(* IEC 61131-3 sources: plcrex/tests/st_examples, 88 files *)

(* ---- TC003.st ---- *)
// ********************************************************************************
// Program Organization Units: FUNCTION
// ********************************************************************************

FUNCTION TC003
  VAR_OUTPUT
    x1 : BOOL;
  END_VAR

  x1 := TRUE;
END_FUNCTION

(* ---- TC004.st ---- *)
// ********************************************************************************
// Program Organization Units: FUNCTION : DATATYPE
// ********************************************************************************

FUNCTION TC004 : BOOL
    VAR_INPUT
        x1 : BOOL;
    END_VAR
    VAR
        x2: BOOL := FALSE;
    END_VAR

    TC004 := x2;
END_FUNCTION

(* ---- TC005.st ---- *)
// ********************************************************************************
// Program Organization Units: FUNCTION_BLOCK
// ********************************************************************************

FUNCTION_BLOCK TC005
  VAR
    x1 : BOOL;
  END_VAR

  x1:= TRUE;
END_FUNCTION_BLOCK

(* ---- TC006.st ---- *)
// ********************************************************************************
// Variable Declaration List: VAR
// ********************************************************************************

FUNCTION_BLOCK TC006
  VAR
    x1 : BOOL := FALSE;
  END_VAR

  x1:= TRUE;
END_FUNCTION_BLOCK

(* ---- TC006_fbd.st ---- *)
FUNCTION_BLOCK TC006
  VAR_INPUT
    i1 : BOOL;
    i2 : BOOL;
  END_VAR
  VAR_OUTPUT
    o1 : BOOL;
    o2 : BOOL;
    o3 : BOOL;
  END_VAR
  VAR
    l1 : BOOL;
    l2 : TIME := T#5s;
    TON0 : TON;
    AND1_OUT : BOOL;
    XOR3_OUT : BOOL;
    OR13_OUT : BOOL;
  END_VAR

  AND1_OUT := AND(i1, i2);
  TON0(AND1_OUT, l2);
  XOR3_OUT := XOR(AND1_OUT, TON0.Q);
  l1 := XOR3_OUT;
  o1 := TON0.Q;
  o2 := i1;
  OR13_OUT := OR(i2, l1);
  o3 := OR13_OUT;
END_FUNCTION_BLOCK

(* ---- TC007.st ---- *)
// ********************************************************************************
// Interface Declaration List: VAR_INPUT
// ********************************************************************************

FUNCTION_BLOCK TC007
  VAR_INPUT
    x1 : BOOL;
  END_VAR
  VAR
    x2 : BOOL := FALSE;
    x3 : BOOL := FALSE;
  END_VAR

  x2:=x1;
END_FUNCTION_BLOCK

(* ---- TC008.st ---- *)
// ********************************************************************************
// Interface Declaration List: VAR_INPUT
// ********************************************************************************

FUNCTION_BLOCK TC008
  VAR_INPUT
    x1 : BOOL := FALSE;
  END_VAR
  VAR
    x2 : BOOL := FALSE;
    x3 : BOOL := FALSE;
  END_VAR

  x2:=x1;
END_FUNCTION_BLOCK

(* ---- TC009.st ---- *)
// ********************************************************************************
// Interface Declaration List: VAR_OUTPUT
// ********************************************************************************

FUNCTION_BLOCK TC009
  VAR_OUTPUT
    x1 : BOOL;
  END_VAR

  x1 := TRUE;
END_FUNCTION_BLOCK

(* ---- TC010.st ---- *)
// ********************************************************************************
// Interface Declaration List: VAR_OUTPUT
// ********************************************************************************

FUNCTION_BLOCK TC010
  VAR_OUTPUT
    x1 : BOOL := FALSE;
  END_VAR

  x1 := TRUE;
END_FUNCTION_BLOCK

(* ---- TC011.st ---- *)
// ********************************************************************************
// Interface Declaration List: VAR_EXTERNAL
// ********************************************************************************

FUNCTION_BLOCK TC011
  VAR_EXTERNAL
    global : BOOL;
  END_VAR
  VAR
    x1 : BOOL;
  END_VAR

  x1 := global;
END_FUNCTION_BLOCK

(* ---- TC012.st ---- *)
// ********************************************************************************
// Interface Declaration List: VAR_IN_OUT
// ********************************************************************************

FUNCTION_BLOCK TC012
  VAR_IN_OUT
    x1 : BOOL;
  END_VAR

  x1:=TRUE;
END_FUNCTION_BLOCK

(* ---- TC013.st ---- *)
// ********************************************************************************
// Data Types: BOOL
// ********************************************************************************

FUNCTION_BLOCK TC013
  VAR
    x1 : BOOL;
  END_VAR

  x1:=TRUE;
END_FUNCTION_BLOCK

(* ---- TC014.st ---- *)
// ********************************************************************************
// Data Types: INT
// ********************************************************************************

FUNCTION_BLOCK TC014
  VAR
    x1 : INT;
  END_VAR

  x1:=5;
END_FUNCTION_BLOCK

(* ---- TC015.st ---- *)
// ********************************************************************************
// Data Types: DINT
// ********************************************************************************

FUNCTION_BLOCK TC015
  VAR
    x1 : DINT;
  END_VAR

  x1:=5;
END_FUNCTION_BLOCK

(* ---- TC016.st ---- *)
// ********************************************************************************
// Data Types: UINT
// ********************************************************************************

FUNCTION_BLOCK TC016
  VAR
    x1 : UINT;
  END_VAR

  x1:=5;
END_FUNCTION_BLOCK

(* ---- TC017.st ---- *)
// ********************************************************************************
// Data Types: REAL
// ********************************************************************************

FUNCTION_BLOCK TC017
  VAR
    x1 : REAL;
  END_VAR

  x1:=5.0;
END_FUNCTION_BLOCK

(* ---- TC018.st ---- *)
// ********************************************************************************
// Data Types: TIME
// ********************************************************************************

FUNCTION_BLOCK TC018
  VAR
    x1 : TIME;
  END_VAR

  x1:=t#5000ms;
END_FUNCTION_BLOCK

(* ---- TC019.st ---- *)
// ********************************************************************************
// Data Types: ARRAY OF BOOL
// ********************************************************************************

FUNCTION_BLOCK TC019
  VAR
    x1 : ARRAY [1..2] OF BOOL;
  END_VAR

  x1[1]:= TRUE;
END_FUNCTION_BLOCK

(* ---- TC020.st ---- *)
// ********************************************************************************
// Data Types: ARRAY OF INT
// ********************************************************************************

FUNCTION_BLOCK TC020
  VAR
    x1 : ARRAY [1..2] OF INT;
  END_VAR

  x1[1]:= 1;
END_FUNCTION_BLOCK

(* ---- TC021.st ---- *)
// ********************************************************************************
// Data Types: ARRAY OF DINT
// ********************************************************************************

FUNCTION_BLOCK TC021
  VAR
    x1 : ARRAY [1..2] OF DINT;
  END_VAR

  x1[1]:= 1;
END_FUNCTION_BLOCK

(* ---- TC022.st ---- *)
// ********************************************************************************
// Data Types: ARRAY OF UINT
// ********************************************************************************

FUNCTION_BLOCK TC022
  VAR
    x1 : ARRAY [1..2] OF UINT;
  END_VAR

  x1[1]:= 1;
END_FUNCTION_BLOCK

(* ---- TC023.st ---- *)
// ********************************************************************************
// Data Types: ARRAY OF REAL
// ********************************************************************************

FUNCTION_BLOCK TC023
  VAR
    x1 : ARRAY [1..2] OF REAL;
  END_VAR

  x1[1]:= 1.0;
END_FUNCTION_BLOCK

(* ---- TC024.st ---- *)
// ********************************************************************************
// Data Types: ARRAY OF TIME
// ********************************************************************************

FUNCTION_BLOCK TC024
  VAR
    x1 : ARRAY [1..2] OF TIME;
  END_VAR

  x1[1]:= t#5000ms;
END_FUNCTION_BLOCK

(* ---- TC025.st ---- *)
// ********************************************************************************
// Expressions: FALSE
// ********************************************************************************

FUNCTION_BLOCK TC025
  VAR
    x1 : BOOL;
  END_VAR

  x1:=FALSE;
END_FUNCTION_BLOCK

(* ---- TC026.st ---- *)
// ********************************************************************************
// Expressions: TRUE
// ********************************************************************************

FUNCTION_BLOCK TC026
  VAR
    x1 : BOOL;
  END_VAR

  x1:=TRUE;
END_FUNCTION_BLOCK

(* ---- TC027.st ---- *)
// ********************************************************************************
// Expressions: =
// ********************************************************************************

FUNCTION_BLOCK TC027
  VAR
    x1 : INT := 4;
    x2 : INT := 6;
    x3 : BOOL;
  END_VAR

  x3:=x1 = x2;
END_FUNCTION_BLOCK

(* ---- TC028.st ---- *)
// ********************************************************************************
// Expressions: =
// ********************************************************************************

FUNCTION_BLOCK TC028
  VAR
    x1 : INT := 6;
    x2 : INT := 6;
    x3 : BOOL;
  END_VAR

  x3:=x1 = x2;
END_FUNCTION_BLOCK

(* ---- TC029.st ---- *)
// ********************************************************************************
// Expressions: <>
// ********************************************************************************

FUNCTION_BLOCK TC029
  VAR
    x1 : INT := 4;
    x2 : INT := 6;
    x3 : BOOL;
  END_VAR

  x3:=x1 <> x2;
END_FUNCTION_BLOCK

(* ---- TC030.st ---- *)
// ********************************************************************************
// Expressions: <>
// ********************************************************************************

FUNCTION_BLOCK TC030
  VAR
    x1 : INT := 6;
    x2 : INT := 6;
    x3 : BOOL;
  END_VAR

  x3:=x1 <> x2;
END_FUNCTION_BLOCK

(* ---- TC031.st ---- *)
// ********************************************************************************
// Expressions: <
// ********************************************************************************

FUNCTION_BLOCK TC031
  VAR
    x1 : INT := 4;
    x2 : INT := 6;
    x3 : BOOL;
  END_VAR

  x3:=x1 < x2;
END_FUNCTION_BLOCK

(* ---- TC032.st ---- *)
// ********************************************************************************
// Expressions: <
// ********************************************************************************

FUNCTION_BLOCK TC032
  VAR
    x1 : INT := 6;
    x2 : INT := 6;
    x3 : BOOL;
  END_VAR

  x3:=x1 < x2;
END_FUNCTION_BLOCK

(* ---- TC033.st ---- *)
// ********************************************************************************
// Expressions: >
// ********************************************************************************

FUNCTION_BLOCK TC033
  VAR
    x1 : INT := 4;
    x2 : INT := 6;
    x3 : BOOL;
  END_VAR

  x3:=x1 > x2;
END_FUNCTION_BLOCK

(* ---- TC034.st ---- *)
// ********************************************************************************
// Expressions: >
// ********************************************************************************

FUNCTION_BLOCK TC034
  VAR
    x1 : INT := 6;
    x2 : INT := 6;
    x3 : BOOL;
  END_VAR

  x3:=x1 > x2;
END_FUNCTION_BLOCK

(* ---- TC035.st ---- *)
// ********************************************************************************
// Expressions: <=
// ********************************************************************************

FUNCTION_BLOCK TC035
  VAR
    x1 : INT := 4;
    x2 : INT := 6;
    x3 : BOOL;
  END_VAR

  x3:=x1 <= x2;
END_FUNCTION_BLOCK

(* ---- TC036.st ---- *)
// ********************************************************************************
// Expressions: <=
// ********************************************************************************

FUNCTION_BLOCK TC036
  VAR
    x1 : INT := 6;
    x2 : INT := 6;
    x3 : BOOL;
  END_VAR

  x3:=x1 <= x2;
END_FUNCTION_BLOCK

(* ---- TC037.st ---- *)
// ********************************************************************************
// Expressions: >=
// ********************************************************************************

FUNCTION_BLOCK TC037
  VAR
    x1 : INT := 4;
    x2 : INT := 6;
    x3 : BOOL;
  END_VAR

  x3:=x1 >= x2;
END_FUNCTION_BLOCK

(* ---- TC038.st ---- *)
// ********************************************************************************
// Expressions: >=
// ********************************************************************************

FUNCTION_BLOCK TC038
  VAR
    x1 : INT := 6;
    x2 : INT := 6;
    x3 : BOOL;
  END_VAR

  x3:=x1 >= x2;
END_FUNCTION_BLOCK

(* ---- TC039.st ---- *)
// ********************************************************************************
// Expressions: NOT
// ********************************************************************************

FUNCTION_BLOCK TC039
  VAR
    x1 : BOOL := TRUE;
    x2 : BOOL;
  END_VAR

  x1:=NOT x1;
  x2 := TRUE;
END_FUNCTION_BLOCK

(* ---- TC040.st ---- *)
// ********************************************************************************
// Expressions: NOT
// ********************************************************************************

FUNCTION_BLOCK TC040
  VAR
    x1 : BOOL := FALSE;
    x2 : BOOL;
  END_VAR

  x1:=NOT x1;
  x2 := TRUE;
END_FUNCTION_BLOCK

(* ---- TC041.st ---- *)
// ********************************************************************************
// Expressions: AND
// ********************************************************************************

FUNCTION_BLOCK TC041
  VAR
    x1 : BOOL := FALSE;
    x2 : BOOL := FALSE;
	x3 : BOOL;
  END_VAR

  x3:=x1 AND x2;
END_FUNCTION_BLOCK

(* ---- TC042.st ---- *)
// ********************************************************************************
// Expressions: AND
// ********************************************************************************

FUNCTION_BLOCK TC042
  VAR
    x1 : BOOL := TRUE;
    x2 : BOOL := FALSE;
	x3 : BOOL;
  END_VAR

  x3:=x1 AND x2;
END_FUNCTION_BLOCK

(* ---- TC043.st ---- *)
// ********************************************************************************
// Expressions: AND
// ********************************************************************************

FUNCTION_BLOCK TC043
  VAR
    x1 : BOOL := FALSE;
    x2 : BOOL := TRUE;
	x3 : BOOL;
  END_VAR

  x3:=x1 AND x2;
END_FUNCTION_BLOCK

(* ---- TC044.st ---- *)
// ********************************************************************************
// Expressions: AND
// ********************************************************************************

FUNCTION_BLOCK TC044
  VAR
    x1 : BOOL := FALSE;
    x2 : BOOL := TRUE;
	x3 : BOOL;
  END_VAR

  x3:=x1 AND x2;
END_FUNCTION_BLOCK

(* ---- TC045.st ---- *)
// ********************************************************************************
// Expressions: XOR
// ********************************************************************************

FUNCTION_BLOCK TC045
  VAR
    x1 : BOOL := FALSE;
    x2 : BOOL := FALSE;
	x3 : BOOL;
  END_VAR

  x3:=x1 XOR x2;
END_FUNCTION_BLOCK

(* ---- TC046.st ---- *)
// ********************************************************************************
// Expressions: XOR
// ********************************************************************************

FUNCTION_BLOCK TC046
  VAR
    x1 : BOOL := TRUE;
    x2 : BOOL := FALSE;
	x3 : BOOL;
  END_VAR

  x3:=x1 XOR x2;
END_FUNCTION_BLOCK

(* ---- TC047.st ---- *)
// ********************************************************************************
// Expressions: XOR
// ********************************************************************************

FUNCTION_BLOCK TC047
  VAR
    x1 : BOOL := FALSE;
    x2 : BOOL := TRUE;
	x3 : BOOL;
  END_VAR

  x3:=x1 XOR x2;
END_FUNCTION_BLOCK

(* ---- TC048.st ---- *)
// ********************************************************************************
// Expressions: XOR
// ********************************************************************************

FUNCTION_BLOCK TC048
  VAR
    x1 : BOOL := TRUE;
    x2 : BOOL := TRUE;
	x3 : BOOL;
  END_VAR

  x3:=x1 XOR x2;
END_FUNCTION_BLOCK

(* ---- TC049.st ---- *)
// ********************************************************************************
// Expressions: OR
// ********************************************************************************

FUNCTION_BLOCK TC049
  VAR
    x1 : BOOL := FALSE;
    x2 : BOOL := FALSE;
	x3 : BOOL;
  END_VAR

  x3:=x1 OR x2;
END_FUNCTION_BLOCK

(* ---- TC050.st ---- *)
// ********************************************************************************
// Expressions: OR
// ********************************************************************************

FUNCTION_BLOCK TC050
  VAR
    x1 : BOOL := TRUE;
    x2 : BOOL := FALSE;
	x3 : BOOL;
  END_VAR

  x3:=x1 OR x2;
END_FUNCTION_BLOCK

(* ---- TC051.st ---- *)
// ********************************************************************************
// Expressions: OR
// ********************************************************************************

FUNCTION_BLOCK TC051
  VAR
    x1 : BOOL := FALSE;
    x2 : BOOL := TRUE;
	x3 : BOOL;
  END_VAR

  x3:=x1 OR x2;
END_FUNCTION_BLOCK

(* ---- TC052.st ---- *)
// ********************************************************************************
// Expressions: OR
// ********************************************************************************

FUNCTION_BLOCK TC052
  VAR
    x1 : BOOL := TRUE;
    x2 : BOOL := TRUE;
	x3 : BOOL;
  END_VAR

  x3:=x1 OR x2;
END_FUNCTION_BLOCK

(* ---- TC053.st ---- *)
// ********************************************************************************
// Expressions: EXPT Macro
// ********************************************************************************

FUNCTION_BLOCK TC053
  VAR
    x1 : REAL := 1.0;
    x2 : REAL := 2.0;
	x3 : REAL;
  END_VAR

  x3:=EXPT(x1,x2);
END_FUNCTION_BLOCK

(* ---- TC054.st ---- *)
// ********************************************************************************
// Expressions: -Tau
// ********************************************************************************

FUNCTION_BLOCK TC054
  VAR
    x1 : INT;
	x2 : INT := 5;
  END_VAR

  x1 := -x2;
END_FUNCTION_BLOCK

(* ---- TC055.st ---- *)
// ********************************************************************************
// Expressions: -Tau
// ********************************************************************************

FUNCTION_BLOCK TC055
  VAR
    x1 : INT;
	x2 : INT := 5;
  END_VAR

  x1 := -(2);
END_FUNCTION_BLOCK

(* ---- TC056.st ---- *)
// ********************************************************************************
// Expressions: *
// ********************************************************************************

FUNCTION_BLOCK TC056
  VAR
    x1 : INT;
    x2 : INT :=5;
  END_VAR

  x1:=x2*3;
END_FUNCTION_BLOCK

(* ---- TC057.st ---- *)
// ********************************************************************************
// Expressions: /
// ********************************************************************************

FUNCTION_BLOCK TC057
  VAR
    x1 : INT;
    x2 : INT :=5;
  END_VAR

  x1:=x2/3;
END_FUNCTION_BLOCK

(* ---- TC058.st ---- *)
// ********************************************************************************
// Expressions: /
// ********************************************************************************

FUNCTION_BLOCK TC058
  VAR
    x1 : REAL;
    x2 : REAL :=5.0;
  END_VAR

  x1:=x2/3.0;
END_FUNCTION_BLOCK

(* ---- TC059.st ---- *)
// ********************************************************************************
// Expressions: MOD
// ********************************************************************************

FUNCTION_BLOCK TC059
  VAR
    x1 : INT;
    x2 : INT :=5;
  END_VAR

  x1:=x2 MOD 3;
END_FUNCTION_BLOCK

(* ---- TC060.st ---- *)
// ********************************************************************************
// Expressions: +
// ********************************************************************************

FUNCTION_BLOCK TC060
  VAR
    x1 : INT;
    x2 : INT :=5;
  END_VAR

  x1:=x2 + 3;
END_FUNCTION_BLOCK

(* ---- TC061.st ---- *)
// ********************************************************************************
// Expressions: -
// ********************************************************************************

FUNCTION_BLOCK TC061
  VAR
    x1 : INT;
    x2 : INT :=5;
  END_VAR

  x1:=x2 - 3;
END_FUNCTION_BLOCK

(* ---- TC062.st ---- *)
// ********************************************************************************
// Expressions: ()
// ********************************************************************************

FUNCTION_BLOCK TC062
  VAR
    x1 : INT;
    x2 : INT :=5;
  END_VAR

  x1:= (1+7) / 3;
END_FUNCTION_BLOCK

(* ---- TC063.st ---- *)
// ********************************************************************************
// Expressions: ()
// ********************************************************************************

FUNCTION_BLOCK TC063
  VAR
    x1 : INT;
    x2 : INT :=5;
  END_VAR

  x1:= (1-7) / 3;
END_FUNCTION_BLOCK

(* ---- TC064.st ---- *)
// ********************************************************************************
// Expressions: ()
// ********************************************************************************

FUNCTION_BLOCK TC064
  VAR
    x1 : REAL;
    x2 : INT :=5;
  END_VAR

  x1:= (1.0-7) / 3.0;
END_FUNCTION_BLOCK

(* ---- TC065.st ---- *)
// ********************************************************************************
// Conditional Statements: IF ELSE
// ********************************************************************************

FUNCTION_BLOCK TC065
  VAR
    x1 : BOOL := TRUE;
    x2 : INT := 5;
	x3 : INT;
  END_VAR

  IF x1 THEN
    x3:=x2;
  END_IF;
END_FUNCTION_BLOCK

(* ---- TC066.st ---- *)
// ********************************************************************************
// Conditional Statements: IF ELSE
// ********************************************************************************

FUNCTION_BLOCK TC066
  VAR
    x1 : BOOL := TRUE;
    x2 : INT := 5;
	x3 : INT;
  END_VAR

  IF x1 THEN
    x3:=x2;
  ELSE
    x3:= -x2;
  END_IF;
END_FUNCTION_BLOCK

(* ---- TC067.st ---- *)
// ********************************************************************************
// Conditional Statements: IF ELSE
// ********************************************************************************

FUNCTION_BLOCK TC067
  VAR
    x1 : BOOL := TRUE;
    x2 : INT := 5;
	x3 : INT;
  END_VAR

  IF x1 THEN
    x3:=x2;
  ELSIF x2 = 5 THEN
    x3:=-x2;
  END_IF;
END_FUNCTION_BLOCK

(* ---- TC068.st ---- *)
// ********************************************************************************
// Conditional Statements: IF ELSE
// ********************************************************************************

FUNCTION_BLOCK TC068
  VAR
    x1 : BOOL := TRUE;
    x2 : INT := 5;
	x3 : INT;
  END_VAR

  IF x1 THEN
    x3:=x2;
  ELSIF x2 = 5 THEN
    x3:=-x2;
  ELSE
    x3:=2*x2;
  END_IF;
END_FUNCTION_BLOCK

(* ---- TC069.st ---- *)
// ********************************************************************************
// Bounded Loops: FOR
// ********************************************************************************

FUNCTION_BLOCK TC069
  VAR
    x1 : INT;
    x2 : INT;
  END_VAR

  FOR x1:=0 TO 10 BY 2 DO
  	x2 := x1+5;
  END_FOR;
END_FUNCTION_BLOCK

(* ---- TC070.st ---- *)
// ********************************************************************************
// Bounded Loops: FOR
// ********************************************************************************

FUNCTION_BLOCK TC070
  VAR
    x2 : INT;
  END_VAR

  FOR x1:=0 TO 10 DO
  	x2 := x1;
  END_FOR;
END_FUNCTION_BLOCK

(* ---- TC071.st ---- *)
// ********************************************************************************
// Bounded Loops: WHILE
// ********************************************************************************

FUNCTION_BLOCK TC071
  VAR
    x1 : INT;
    x2 : INT;
  END_VAR

  WHILE x1 <= 10 DO
  	x1 := x2 + x1;
  END_WHILE;
END_FUNCTION_BLOCK

(* ---- TC072.st ---- *)
// ********************************************************************************
// Bounded Loops: REPEAT UNTIL
// ********************************************************************************

FUNCTION_BLOCK TC072
  VAR
    x1 : INT;
    x2 : INT;
  END_VAR

  REPEAT
  	x1 := 5 + x2;
  UNTIL x1 > 10
  END_REPEAT;
END_FUNCTION_BLOCK

(* ---- TC073.st ---- *)
// ********************************************************************************
// Assignment: :=
// ********************************************************************************

FUNCTION_BLOCK TC073
  VAR
    x1 : INT;
    x2 : INT;
    x3 : INT;
  END_VAR

  x1:=1;
  x2:=1;
  x3:=1;

END_FUNCTION_BLOCK

(* ---- TC074.st ---- *)
// ********************************************************************************
// Assignment: :=
// ********************************************************************************

FUNCTION_BLOCK TC074
  VAR
    x1 : INT;
    x2 : INT;
    x3 : INT;
  END_VAR

  x1:=1;
  x2:=1;
  x1:=2;

END_FUNCTION_BLOCK

(* ---- TC075.st ---- *)
// ********************************************************************************
// Assignment: :=
// ********************************************************************************

FUNCTION_BLOCK TC075
  VAR
    x1 : INT;
    x2 : INT;
    x3 : INT;
  END_VAR

  x1:=x1+2;
  x2:=1;

END_FUNCTION_BLOCK

(* ---- TC076.st ---- *)
// ********************************************************************************
// Assignment: :=
// ********************************************************************************

FUNCTION_BLOCK TC076
  VAR
    x1 : INT;
    x2 : INT;
    x3 : INT;
  END_VAR

  x1:=2;
  x1:=3;

END_FUNCTION_BLOCK

(* ---- TC077.st ---- *)
// ********************************************************************************
// Assignment: :=
// ********************************************************************************

FUNCTION_BLOCK TC077
  VAR
    x1 : INT;
    x2 : INT;
    x3 : INT;
  END_VAR

  x1:=x2;
  x2:=1;

END_FUNCTION_BLOCK

(* ---- TC078.st ---- *)
// ********************************************************************************
// Assignment: :=
// ********************************************************************************

FUNCTION_BLOCK TC078
  VAR
    x1 : INT;
    x2 : INT;
    x3 : INT;
  END_VAR

  x1:=1;
  x2:=x1;

END_FUNCTION_BLOCK

(* ---- TC079.st ---- *)
// ********************************************************************************
// Assignment: :=
// ********************************************************************************

FUNCTION_BLOCK TC079
  VAR
    x1 : INT;
    x2 : INT;
    x3 : INT;
  END_VAR

  x1:=x1+1;

END_FUNCTION_BLOCK

(* ---- TC080.st ---- *)
// ********************************************************************************
// Real POU
// ********************************************************************************

FUNCTION_BLOCK TC080
	VAR_INPUT
		S1 : BOOL;
		R : BOOL;
	END_VAR
	VAR_OUTPUT
		Q1 : BOOL;
	END_VAR

	Q1 := S1 XOR (Q1 AND NOT R);
END_FUNCTION_BLOCK

(* ---- TC081.st ---- *)
FUNCTION_BLOCK TC081
	VAR_INPUT
		IN1 : INT;
		IN2 : INT;
		IN3 : INT;
		IN4 : BOOL;
	END_VAR
	VAR_OUTPUT
		Wrn : BOOL;
		Err : BOOL;
		Ctr : INT;
		iOut2 : INT;
	END_VAR
	VAR
	    SR1 : SR;
	    TON1 : TON;
	    TON2 : TON;
	END_VAR

    SR1(((((20*IN1)+(6*IN2)+IN3))=(100*2)) AND (IN1+IN2+IN3=100),IN4);
    TON1((((((20*IN1)+(6*IN2)+IN3))=(100*2)) AND (IN1+IN2+IN3=100)),2);
    TON2(IN1+IN2+IN3=42 AND SR1.Q,3);
    Ctr := TON2.ET;
    Err := TON1.Q;
    Wrn := SR1.Q;
END_FUNCTION_BLOCK

(* ---- TC082.st ---- *)
// ********************************************************************************
// Real POU
// ********************************************************************************

FUNCTION_BLOCK TC082
  VAR_INPUT
    IN : BOOL;
	PT : INT;
  END_VAR
  VAR_OUTPUT
    Q : BOOL;
	ET : INT;
  END_VAR
  VAR
    CYCLE : INT;
    TIMER : INT;
    TIMERN : INT;
    GE7_OUT : BOOL;
    ADD8_OUT : INT;
    SEL3_OUT : INT;
    SEL5_OUT : INT;
    SEL2_OUT : INT;
    SEL6_OUT : INT;
    SEL1_OUT : BOOL;
    SEL4_OUT : BOOL;
  END_VAR

  GE7_OUT := GE(TIMER, PT);
  ADD8_OUT := ADD(TIMER, CYCLE);
  SEL3_OUT := SEL(GE7_OUT, TIMER, ADD8_OUT);
  SEL5_OUT := SEL(IN, SEL3_OUT, 0);
  SEL2_OUT := SEL(GE7_OUT, PT, TIMER);
  SEL6_OUT := SEL(IN, SEL2_OUT, 0);
  SEL1_OUT := SEL(GE7_OUT, true, false);
  SEL4_OUT := SEL(IN, SEL1_OUT, false);
  Q := SEL4_OUT;
  ET := SEL6_OUT;
  TIMERN := SEL5_OUT;
  TIMER := TIMERN;
END_FUNCTION_BLOCK

(* ---- _TC001.st ---- *)
 PROGRAM TC001
 VAR_INPUT
 x1:INT;
 END_VAR
 VAR_OUTPUT
 x2:INT;
 END_VAR
 VAR
 x3:INT:=3;
 END_VAR
 x2:=x1+x3;
 END_PROGRAM

(* ---- TC001.st ---- *)
// ********************************************************************************
// Program Organization Units: PROGRAM
// ********************************************************************************

PROGRAM TC001
  VAR_INPUT
    x1 : INT;
  END_VAR
  VAR_OUTPUT
    x2 : INT;
  END_VAR
  VAR
    x3 : INT := 3;
  END_VAR

  x2:=x1+x3;
END_PROGRAM

(* ---- TC002.st ---- *)
// ********************************************************************************
// Program Organization Units: PROGRAM
// ********************************************************************************

PROGRAM TC002
  VAR_INPUT
    x1 : INT;
  END_VAR
  VAR_OUTPUT
    x2 : INT;
  END_VAR
  VAR
    x3 : INT := 3;
  END_VAR

  x2:=x1 +(x3*x1);
END_PROGRAM

(* ---- TC005_fbd.st ---- *)
PROGRAM TC005
        VAR_INPUT
                i1 : BOOL;
                i2 : BOOL := FALSE;
                i3 : TIME;
        END_VAR
        VAR_OUTPUT
                o1 : BOOL := FALSE;
                o2 : BOOL := FALSE;
        END_VAR
        VAR
                o4 : BOOL;
                TON0 : TON;
                AND1_OUT : BOOL;
                XOR3_OUT : BOOL;
        END_VAR

        AND1_OUT := AND(i1,i2);
        TON0(AND1_OUT,i3);
        XOR3_OUT := XOR(AND1_OUT,TON0.Q);
        o1 := XOR3_OUT;
        o4 := TON0.Q;
        o2 := i1;
END_PROGRAM

(* ---- TC083.st ---- *)
PROGRAM TC083
  VAR_ACCESS
    Var1 : DINT;
    Var2 : DINT;
    Var3 : DINT;
  END_VAR

  Var1 := 19 / 0;
  Var2 := Var1 / 1;
END_PROGRAM

(* ---- TC084.st ---- *)
FUNCTION dead_code_after_return : INT
  VAR
    counter : INT := 0;
    some_var : INT;
  END_VAR
  counter := counter + 1;
  counter := 2 + 2;
  RETURN;
  some_var := SQRT(16#42); (* UnreachableCode error *)
  some_var := 16#42; (* No additional warnings *)
  some_var := 19;
END_FUNCTION

PROGRAM dead_code_in_the_loops
VAR a : INT; i : INT; END_VAR
  WHILE i < 10 DO
    IF i = 5 THEN
      i := i + 1;
      EXIT;
      i := 19; (* UnreachableCode error *)
      i := 42; (* No additional warnings *)
      i := 42;
    ELSIF i = 6 THEN
      CONTINUE;
      i := 3; (* UnreachableCode error *)
      i := 44; (* No additional warnings *)
      i := 19;
    END_IF;
    i := i + 2;
  END_WHILE;
  I := 0;
END_PROGRAM

(* ---- TC085.st ---- *)
PROGRAM TC085
  VAR_INPUT
    a: INT;
    b: INT;
  END_VAR
  VAR_OUTPUT
    gcd:INT;
  END_VAR
  VAR
    c: INT;
    d: INT;
  END_VAR

    c:=a;
    d:=b;

    IF (c=0) THEN
        gcd := d;

    ELSE
        WHILE (d <>0) DO
            IF (c>d) THEN
                c := c-d;
            ELSE
                d := d-c;
            END_IF;
        END_WHILE;
        gcd := c;
    END_IF;
END_PROGRAM
